(* IEC 61131-3 sources: IRIS-Project/LASAL CONTROL SOFTWARE/LasalProject_2025_09_12/Class/ExactStep, 1 file *)

(* ---- ExactStep.st ---- *)
(*!
<Class
	Name               = "ExactStep"
	Revision           = "0.0"
	RealtimeTask       = "false"
	CyclicTask         = "true"
	DefCyclictime      = "200 ms"
	BackgroundTask     = "false"
	Sigmatek           = "false"
	OSInterface        = "false"
	HighPriority       = "false"
	Automatic          = "false"
	UpdateMode         = "Prescan"
	SharedCommandTable = "true"
	Objectsize         = "(574,120)">
	<Channels>
		<Server Name="ClassSvr" Visualized="false" Initialize="false" WriteProtected="true" Retentive="false"/>
		<Server Name="M1_EXACT_STEP" Visualized="false" Initialize="false" WriteProtected="false" Retentive="false"/>
		<Server Name="M3_EXACT_STEP" Visualized="false" Initialize="false" WriteProtected="false" Retentive="false"/>
		<Server Name="M4_EXACT_STEP" Visualized="false" Initialize="false" WriteProtected="false" Retentive="false"/>
		<Server Name="M5_EXACT_CS_1" Visualized="false" Initialize="false" WriteProtected="false" Retentive="false"/>
		<Server Name="M5_EXACT_CS_2" Visualized="false" Initialize="false" WriteProtected="false" Retentive="false"/>
		<Server Name="M5_EXACT_CS_3" Visualized="false" Initialize="false" WriteProtected="false" Retentive="false"/>
		<Server Name="M5_EXACT_DS" Visualized="false" Initialize="false" WriteProtected="false" Retentive="false"/>
		<Server Name="M5_EXACT_IS_1" Visualized="false" Initialize="false" WriteProtected="false" Retentive="false"/>
		<Server Name="M5_EXACT_IS_2" Visualized="false" Initialize="false" WriteProtected="false" Retentive="false"/>
		<Server Name="M5_EXACT_IS_3" Visualized="false" Initialize="false" WriteProtected="false" Retentive="false"/>
		<Server Name="M5_OFFSET_DS" Visualized="false" Initialize="false" WriteProtected="false" Retentive="false"/>
	</Channels>
</Class>
*)
ExactStep : CLASS
  //Servers:
	ClassSvr 	: SvrChCmd_DINT;
	M1_EXACT_STEP 	: SvrCh_DINT;
	M3_EXACT_STEP 	: SvrCh_DINT;
	M4_EXACT_STEP 	: SvrCh_DINT;
	M5_EXACT_CS_1 	: SvrCh_DINT;
	M5_EXACT_CS_2 	: SvrCh_DINT;
	M5_EXACT_CS_3 	: SvrCh_DINT;
	M5_EXACT_IS_1 	: SvrCh_DINT;
	M5_EXACT_IS_2 	: SvrCh_DINT;
	M5_EXACT_IS_3 	: SvrCh_DINT;
	M5_EXACT_DS 	: SvrCh_DINT;
	M5_OFFSET_DS 	: SvrCh_DINT;
  //Clients:
  //Variables:
  //Functions:

	FUNCTION VIRTUAL GLOBAL CyWork
		VAR_INPUT
			EAX 	: UDINT;
		END_VAR
		VAR_OUTPUT
			state (EAX) 	: UDINT;
		END_VAR;

	FUNCTION VIRTUAL GLOBAL Background
		VAR_INPUT
			EAX 	: UDINT;
		END_VAR
		VAR_OUTPUT
			state (EAX) 	: UDINT;
		END_VAR;

	FUNCTION VIRTUAL GLOBAL M1_EXACT_STEP::Read
		VAR_OUTPUT
			output (EAX) 	: DINT;
		END_VAR;

	FUNCTION VIRTUAL GLOBAL M3_EXACT_STEP::Read
		VAR_OUTPUT
			output (EAX) 	: DINT;
		END_VAR;

	FUNCTION VIRTUAL GLOBAL M4_EXACT_STEP::Read
		VAR_OUTPUT
			output (EAX) 	: DINT;
		END_VAR;

	FUNCTION VIRTUAL GLOBAL M5_EXACT_CS_1::Read
		VAR_OUTPUT
			output (EAX) 	: DINT;
		END_VAR;

	FUNCTION VIRTUAL GLOBAL M5_EXACT_CS_2::Read
		VAR_OUTPUT
			output (EAX) 	: DINT;
		END_VAR;

	FUNCTION VIRTUAL GLOBAL M5_EXACT_CS_3::Read
		VAR_OUTPUT
			output (EAX) 	: DINT;
		END_VAR;

	FUNCTION VIRTUAL GLOBAL M5_EXACT_IS_1::Read
		VAR_OUTPUT
			output (EAX) 	: DINT;
		END_VAR;

	FUNCTION VIRTUAL GLOBAL M5_EXACT_IS_2::Read
		VAR_OUTPUT
			output (EAX) 	: DINT;
		END_VAR;

	FUNCTION VIRTUAL GLOBAL M5_EXACT_IS_3::Read
		VAR_OUTPUT
			output (EAX) 	: DINT;
		END_VAR;

	FUNCTION VIRTUAL GLOBAL M5_EXACT_DS::Read
		VAR_OUTPUT
			output (EAX) 	: DINT;
		END_VAR;

	FUNCTION VIRTUAL GLOBAL M5_OFFSET_DS::Read
		VAR_OUTPUT
			output (EAX) 	: DINT;
		END_VAR;
  //Tables:
	FUNCTION @STD
		VAR_OUTPUT
			ret_code	: CONFSTATES;
		END_VAR;
	FUNCTION GLOBAL TAB @CT_;
END_CLASS;

FUNCTION VIRTUAL GLOBAL ExactStep::Background
	VAR_INPUT
		EAX 	: UDINT;
	END_VAR
	VAR_OUTPUT
		state (EAX) 	: UDINT;
	END_VAR

	state := READY;

END_FUNCTION

FUNCTION VIRTUAL GLOBAL ExactStep::M1_EXACT_STEP::Read
	VAR_OUTPUT
		output (EAX) 	: DINT;
	END_VAR

	output := M1_EXACT_STEP;

END_FUNCTION

FUNCTION VIRTUAL GLOBAL ExactStep::M3_EXACT_STEP::Read
	VAR_OUTPUT
		output (EAX) 	: DINT;
	END_VAR

	output := M3_EXACT_STEP;

END_FUNCTION

FUNCTION VIRTUAL GLOBAL ExactStep::M4_EXACT_STEP::Read
	VAR_OUTPUT
		output (EAX) 	: DINT;
	END_VAR

	output := M4_EXACT_STEP;

END_FUNCTION

FUNCTION VIRTUAL GLOBAL ExactStep::M5_EXACT_CS_1::Read
	VAR_OUTPUT
		output (EAX) 	: DINT;
	END_VAR

	output := M5_EXACT_CS_1;

END_FUNCTION

FUNCTION VIRTUAL GLOBAL ExactStep::M5_EXACT_CS_2::Read
	VAR_OUTPUT
		output (EAX) 	: DINT;
	END_VAR

	output := M5_EXACT_CS_2;

END_FUNCTION

FUNCTION VIRTUAL GLOBAL ExactStep::M5_EXACT_CS_3::Read
	VAR_OUTPUT
		output (EAX) 	: DINT;
	END_VAR

	output := M5_EXACT_CS_3;

END_FUNCTION

FUNCTION VIRTUAL GLOBAL ExactStep::M5_EXACT_IS_1::Read
	VAR_OUTPUT
		output (EAX) 	: DINT;
	END_VAR

	output := M5_EXACT_IS_1;

END_FUNCTION

FUNCTION VIRTUAL GLOBAL ExactStep::M5_EXACT_IS_2::Read
	VAR_OUTPUT
		output (EAX) 	: DINT;
	END_VAR

	output := M5_EXACT_IS_2;

END_FUNCTION

FUNCTION VIRTUAL GLOBAL ExactStep::M5_EXACT_IS_3::Read
	VAR_OUTPUT
		output (EAX) 	: DINT;
	END_VAR

	output := M5_EXACT_IS_3;

END_FUNCTION

FUNCTION VIRTUAL GLOBAL ExactStep::M5_EXACT_DS::Read
	VAR_OUTPUT
		output (EAX) 	: DINT;
	END_VAR

	output := M5_EXACT_DS;

END_FUNCTION

FUNCTION VIRTUAL GLOBAL ExactStep::M5_OFFSET_DS::Read
	VAR_OUTPUT
		output (EAX) 	: DINT;
	END_VAR

	output := M5_OFFSET_DS;

END_FUNCTION

FUNCTION VIRTUAL GLOBAL ExactStep::CyWork
	VAR_INPUT
		EAX 	: UDINT;
	END_VAR
	VAR_OUTPUT
		state (EAX) 	: UDINT;
	END_VAR
M1_EXACT_STEP.Write(input:=P_M1_C);
M3_EXACT_STEP.Write(input:=P_M3_C);
M4_EXACT_STEP.Write(input:=P1_M4);

M5_EXACT_CS_1.Write(input:=P1_M5);
M5_EXACT_CS_2.Write(input:=P2_M5);
M5_EXACT_CS_3.Write(input:=P3_M5);

M5_EXACT_IS_1.Write(input:=P1_M5_I);
M5_EXACT_IS_2.Write(input:=P2_M5_I);
M5_EXACT_IS_3.Write(input:=P3_M5_I);

M5_EXACT_DS.Write(input:=P_M5_D);
M5_OFFSET_DS.Write(input:=OffsetDischarge);
	state := READY;

END_FUNCTION
